// TIA Portal V19 export
TYPE "ST_Move"
   STRUCT
      Execute : Bool;
      Distance : Int;
      Velocity : Int;
      Busy : Bool;
      Done : Bool;
      Error : Bool;
      ErrorID : Word;
      CommandAborted : Bool;
   END_STRUCT;
END_TYPE
